(* CODESYS project PLC.project
   Title: 3D_PRINT_TITAN1
   Version: 0.0.0.0

Project tree, tasks and I/O mapping:
  Controller_2A1 : TM241CE24T/U, Schneider Electric, order no. TM241CE24T/U, version 4.0.6.18
    application Application
      libraries: SysTime, 3.4.1.20 (System)
      task MAST (cyclic, interval t#10ms, priority 1, watchdog 1000 ms x 1) calls AVC, Main
      program Main [ST]
      trace Trace_2 (task MAST): Freq_WF1, Freq_WF2, Freq_WF3
      program Wire_Speed_Correction [ST]
      program Manual [ST]
      program Auto [ST]
      trace Trace_3 (task MAST): Process_Auto, MW6, MW4
      program Alarms_manual [ST]
      program Measure [ST]
      trace Trace (task MAST): qiModule_4A1_QW0
      program Alarms_auto [ST]
      trace Trace_1 (task MAST): EM_L_PWM, EM_R_PWM
      program AVC [ST]
      global variables GVL
    Counters : Counters, Schneider Electric, version 4.0.6.18
        settings: A input History = 'old=4 new=-1'; A input History = 'old=4 new=-1'; Instance name = 'HSC0'; A input History = 'old=-1 new=4'; Temporary Instance name = 'HSC0'; Instance name = 'HSC1'; A input History = 'old=-1 new=5'; Temporary Instance name = 'HSC1'; Instance name = 'HSC2'; A input History = 'old=-1 new=6'; Temporary Instance name = 'HSC2'
    Cartridge_1 : Cartridge, Schneider Electric, version 4.0.6.18
    Serial_Line_1 : Serial line, Schneider Electric, version 4.0.6.18
      Modbus_IOScanner : Modbus IOScanner, Schneider Electric, version 3.5.3.8
          settings: Transmission = 'RTU'; ResponseTimeout = 1000; TimeBetweenFrames = 10
        Generic_Modbus_Slave : Generic Modbus Slave, Schneider Electric, version 3.5.3.9
            settings: SlaveAddress = 10; ResponseTimeout = 5000; Output.Function Code = 16; Output.Read Offset = 0; Output.Read Length = 0; Output.Write Offset = 16#0000; Output.Write Length = 1; Output.Cycle Time = 10
            unmapped channels: Output
    DI : Digital Inputs, Schneider Electric, version 4.0.6.18
        settings: IOs Usage = 112
        input  ibDI_IB1 : BYTE  // IB1
        unmapped channels: IW0
    Pulse_Generators : Pulse Generators, Schneider Electric, version 4.0.6.18
        settings: A output History = 'old=0 new=-1'; A output History = 'old=1 new=-1'; A output History = 'old=2 new=-1'
    Serial_Line_2 : Serial line, Schneider Electric, version 4.0.6.18
      Modbus_Manager : Modbus Manager, Schneider Electric, version 4.0.0.2
    DQ : Digital Outputs, Schneider Electric, version 4.0.6.18
        output qwDQ_QW0 : WORD  // QW0
        output qbDQ_QB1 : BYTE  // QB1
    COM_Bus : COM bus, Schneider Electric, version 4.0.6.18
    IO_Bus : IO bus - TM3, Schneider Electric, version 4.0.6.18
      Module_7A1 : TM3AM6/G, Schneider Electric, order no. TM3AM6/G, version 1.0.0.14
          settings: KPI Configuration.KPI Configuration[32] = 19; KPI Configuration.KPI Configuration[33] = 19; KPI Configuration.KPI Configuration[34] = 160; KPI Configuration.KPI Configuration[35] = 15; KPI Configuration.KPI Configuration[36] = 160; KPI Configuration.KPI Configuration[37] = 15; KPI Configuration.KPI Configuration[38] = 32; KPI Configuration.KPI Configuration[39] = 78; KPI Configuration.KPI Configuration[40] = 32; KPI Configuration.KPI Configuration[41] = 78
          input  iiModule_2_IW0 : INT  // IW0
          input  iiModule_2_IW1 : INT  // IW1
          input  iiModule_2_IW2 : INT  // IW2
          input  iiModule_2_IW3 : INT  // IW3
          output qiModule_2_QW0 : INT  // QW0
          output qiModule_2_QW1 : INT  // QW1
          input  ibModule_2_IBStatusIW0 : BYTE  // IBStatusIW0
          input  ibModule_2_IBStatusIW1 : BYTE  // IBStatusIW1
          input  ibModule_2_IBStatusIW2 : BYTE  // IBStatusIW2
          input  ibModule_2_IBStatusIW3 : BYTE  // IBStatusIW3
          input  ibModule_2_IBStatusQW0 : BYTE  // IBStatusQW0
          input  ibModule_2_IBStatusQW1 : BYTE  // IBStatusQW1
      Module_5A1 : TM3AQ4/G, Schneider Electric, order no. TM3AQ4/G, version 1.0.0.12
          settings: KPI Configuration.KPI Configuration[0] = 19; KPI Configuration.KPI Configuration[1] = 19; KPI Configuration.KPI Configuration[2] = 19; KPI Configuration.KPI Configuration[3] = 19; KPI Configuration.KPI Configuration[4] = 160; KPI Configuration.KPI Configuration[5] = 15; KPI Configuration.KPI Configuration[6] = 160; KPI Configuration.KPI Configuration[7] = 15; KPI Configuration.KPI Configuration[8] = 160; KPI Configuration.KPI Configuration[9] = 15; KPI Configuration.KPI Configuration[10] = 160; KPI Configuration.KPI Configuration[11] = 15; KPI Configuration.KPI Configuration[12] = 32; KPI Configuration.KPI Configuration[13] = 78; KPI Configuration.KPI Configuration[14] = 32; KPI Configuration.KPI Configuration[15] = 78; KPI Configuration.KPI Configuration[16] = 32; KPI Configuration.KPI Configuration[17] = 78; KPI Configuration.KPI Configuration[18] = 32; KPI Configuration.KPI Configuration[19] = 78
          output qiModule_5A1_QW0 : INT  // QW0
          output qiModule_5A1_QW1 : INT  // QW1
          output qiModule_5A1_QW2 : INT  // QW2
          output qiModule_5A1_QW3 : INT  // QW3
          input  ibModule_5A1_IBStatusQW0 : BYTE  // IBStatusQW0
          input  ibModule_5A1_IBStatusQW1 : BYTE  // IBStatusQW1
          input  ibModule_5A1_IBStatusQW2 : BYTE  // IBStatusQW2
          input  ibModule_5A1_IBStatusQW3 : BYTE  // IBStatusQW3
      Module_9A1 : TM3TI4/G, Schneider Electric, order no. TM3TI4/G, version 1.0.1.5
          settings: KPI Configuration.KPI Configuration[1] = 35; KPI Configuration.KPI Configuration[2] = 35; KPI Configuration.KPI Configuration[7] = 0; KPI Configuration.KPI Configuration[8] = 160; KPI Configuration.KPI Configuration[9] = 15; KPI Configuration.KPI Configuration[14] = 48; KPI Configuration.KPI Configuration[15] = 117; KPI Configuration.KPI Configuration[16] = 32; KPI Configuration.KPI Configuration[17] = 78; KPI Configuration.KPI Configuration[22] = 5; KPI Configuration.KPI Configuration[24] = 10
          input  iiModule_3_IW0 : INT  // IW0
          input  iiModule_3_IW1 : INT  // IW1
          input  iiModule_3_IW2 : INT  // IW2
          input  iiModule_3_IW3 : INT  // IW3
          input  ibModule_3_IBStatusIW0 : BYTE  // IBStatusIW0
          input  ibModule_3_IBStatusIW1 : BYTE  // IBStatusIW1
          input  ibModule_3_IBStatusIW2 : BYTE  // IBStatusIW2
          input  ibModule_3_IBStatusIW3 : BYTE  // IBStatusIW3
      Module_3A1 : TM3DQ8T/G, Schneider Electric, order no. TM3DQ8T/G, version 1.0.1.4
          output qbModule_1_QB0 : BYTE  // QB0
      Module_3A2 : TM3DQ16R/G, Schneider Electric, order no. TM3DQ16R/G, version 1.0.1.4
          output qwModule_1_QW0 : WORD  // QW0
      Module_4A1 : TM3AQ4/G, Schneider Electric, order no. TM3AQ4/G, version 1.0.0.12
          settings: KPI Configuration.KPI Configuration[0] = 19; KPI Configuration.KPI Configuration[1] = 19; KPI Configuration.KPI Configuration[2] = 19; KPI Configuration.KPI Configuration[3] = 19; KPI Configuration.KPI Configuration[4] = 160; KPI Configuration.KPI Configuration[5] = 15; KPI Configuration.KPI Configuration[6] = 160; KPI Configuration.KPI Configuration[7] = 15; KPI Configuration.KPI Configuration[8] = 160; KPI Configuration.KPI Configuration[9] = 15; KPI Configuration.KPI Configuration[10] = 160; KPI Configuration.KPI Configuration[11] = 15; KPI Configuration.KPI Configuration[12] = 32; KPI Configuration.KPI Configuration[13] = 78; KPI Configuration.KPI Configuration[14] = 32; KPI Configuration.KPI Configuration[15] = 78; KPI Configuration.KPI Configuration[16] = 32; KPI Configuration.KPI Configuration[17] = 78; KPI Configuration.KPI Configuration[18] = 32; KPI Configuration.KPI Configuration[19] = 78
          output qiModule_4A1_QW0 : INT  // QW0
          output qiModule_4A1_QW1 : INT  // QW1
          output qiModule_4A1_QW2 : INT  // QW2
          output qiModule_4A1_QW3 : INT  // QW3
          input  ibModule_4A1_IBStatusQW0 : BYTE  // IBStatusQW0
          input  ibModule_4A1_IBStatusQW1 : BYTE  // IBStatusQW1
          input  ibModule_4A1_IBStatusQW2 : BYTE  // IBStatusQW2
          input  ibModule_4A1_IBStatusQW3 : BYTE  // IBStatusQW3
    Ethernet_Slave : Ethernet Network, Schneider Electric, version 4.0.6.18
        settings: IPAddress = [192, 168, 137, 2]; SubnetMask = [255, 255, 255, 0]; DeviceName = 'PLC_Slave'; WebServer = FALSE; FTP Server = FALSE; SoMachine Protocol = TRUE; Modbus Server = TRUE; NetManage Protocol = FALSE; SNMP protocol = FALSE
  FdtConnections : FDT Connections, Schneider Electric, version 1.0.0.2
    Modbus_Serial_Line_Manager : Modbus Serial Line Manager, Schneider Electric, version 2.2.5
*)

// Controller_2A1/Application/GVL
VAR_GLOBAL
	IX07 AT %IX0.7: BOOL;
	IW19 AT %IW19: WORD ;
	QW13 AT %QW13: WORD;
    Robot_MeasureCmd : BOOL; // 1 = міряти, 0 = зупинити
    Robot_MeasureCmd_Prev : BOOL := FALSE; // Попередній стан сигналу
    // Події
    StartEvent : BOOL := FALSE;
    StopEvent : BOOL := FALSE;
    // Стан вимірювання
    Measuring : BOOL := FALSE;
    MeasureDone : BOOL := FALSE;
    MeasureStatus : INT := 0;     // 0=idle, 1=measuring, 2=done, 3=error
    // Аналоговий сигнал
    VoltageRaw : REAL;
    VoltageFiltered : REAL;
    // Фільтрація
    K_Filter : REAL := 0.12;
    FirstSample : BOOL := TRUE;
    // Обмеження допустимого діапазону
    VoltageMin : REAL := 10.0;
    VoltageMax : REAL := 30.0;
    // Захист від різких викидів
    MaxJump : REAL := 10.0;
    SampleValid : BOOL := FALSE;
    // Накопичення середнього
    VoltageSum : REAL := 0.0;
    SampleCount : DINT := 0;
    VoltageAverage : REAL := 0.0;
    // Результат для Modbus
    VoltageAverage_x100 : WORD := 0;
	
	AVC_ON: BOOL;	
	AVC_Correction AT %QW13: UINT;
	PilotArcIN AT %IX0.0: BOOL;
	PilotArc: BOOL;
	MainArc AT %IX0.1: BOOL;
	//EncoderWF1 AT %IX0.4: BOOL;
	//EncoderWF2 AT %IX0.5: BOOL;
	//EncoderWF3 AT %IX0.6: BOOL;
	StartExt AT %IX1.0: BOOL;
	ReadyExt AT %IX1.1: BOOL;
	EmergencyExt AT %IX1.2: BOOL;
	
	EM_R_PWM AT %QX0.0: BOOL;
	EM_L_PWM AT %QX0.1: BOOL;
	EM_R_EN AT %QX0.2: BOOL;
	EM_L_EN AT %QX0.3: BOOL;
	StartParc AT %QX0.4: BOOL;
	StartMArc AT %QX0.5: BOOL;
	PArcON AT %QX0.6: BOOL;
	ProcON AT %QX0.7: BOOL;
	
	MF1_CW AT %QX3.0: BOOL;
	MF1_CCW AT %QX3.1: BOOL;
	MF2_CW AT %QX3.2: BOOL;
	MF2_CCW AT %QX3.3: BOOL;
	MF3_CW AT %QX3.4: BOOL;
	MF3_CCW AT %QX3.5: BOOL;
	
	Y1 AT %QX4.0: BOOL;
	Y2 AT %QX4.1: BOOL;
	Y3 AT %QX4.2: BOOL;
	Y4 AT %QX4.3: BOOL;
	Y5 AT %QX4.4: BOOL;
	Y6 AT %QX4.5: BOOL;
	Y7 AT %QX4.6: BOOL;
	Y8 AT %QX4.7: BOOL;
	
	PF1 AT %QX5.0: BOOL;
	PF2 AT %QX5.1: BOOL;
	PF3 AT %QX5.2: BOOL;
	PF4 AT %QX5.3: BOOL;
	
	CMT_PS AT %QX5.4: BOOL;
	CMT_PlusI AT %QX5.5: BOOL;
	CMT_MinusI AT %QX5.6: BOOL;
	
	PF1_SPD AT %QW3: WORD;
	PF2_SPD AT %QW4: WORD;
	PF3_SPD AT %QW5: WORD;
	PF4_SPD AT %QW6: WORD;
	
	WF1_SPD AT %QW7: WORD;
	WF2_SPD AT %QW8: WORD;
	WF3_SPD AT %QW9: WORD;
	
	SetCurrent AT %QW11: WORD;
	MeasureU AT %IW14: WORD;
	MeasureI AT %IW15: WORD;
	MeasureU_MHI AT %MW100: WORD;
	MeasureI_MHI AT %MW102: WORD;
	Alarms AT %MW104 : WORD;
	ErrorInManual AT %MW106: WORD;
	
	EmagFreqCalc: REAL;
	Toggle_Ready : BOOL;
	ToggleState : BOOL;
	LastToggleTime : ULINT := 0;
	CurrentTime : ULINT;
    HalfPeriod_us : ULINT;
	
	
	EmagFreqCalc_Auto: REAL;

	Freq_WF1 : REAL := 0.0;
	Freq_WF2 : REAL := 0.0;
	Freq_WF3 : REAL := 0.0;
	Correction : BOOL;
	
	Enable_Start : BOOL;
	
	TON_Delay_Start_PF : TON;
	TON_Delay_Start_WF : TON;
	TON_Delay_Start_Emagnet : TON;
	TON_preblow : TON;
	
	
	MW0 AT %MW0: WORD;
	MW2 AT %MW2: WORD;
	MW4 AT %MW4 : WORD;
	MW6 AT %MW6 : WORD;
	MW8 AT %MW8 : WORD;
	PrevCurrentCMT_HMI : WORD;
END_VAR

VAR_GLOBAL RETAIN	
	EmagFreqSet AT %MD11: REAL;
	
	AVC_Voltage AT %MW12: WORD;
	AVC_Accuracy AT %MW14: WORD;
	AVC_PID_Kp AT %MD8: REAL;
	AVC_PID_Ki AT %MD55: REAL;
	AVC_DELAY AT %MW114: WORD;
	
	SetCurrent_HMI_Man AT %MW20: WORD;
	WF1_SPD_HMI_Man AT %MW26: WORD;
	WF2_SPD_HMI_Man AT %MW28: WORD;
	WF3_SPD_HMI_Man AT %MW30: WORD;
	PF1_SPD_HMI_Man AT %MW32: WORD;
	PF2_SPD_HMI_Man AT %MW34: WORD;
	PF3_SPD_HMI_Man AT %MW36: WORD;
	PF4_SPD_HMI_Man AT %MW38: WORD;
	SetCurrentCMT_HMI AT %MW40: WORD;
	Check_Voltage_Current_Delay AT %MW42 : WORD;
	Emergency_Delay AT %MW44 : WORD;
	Auto_Button_State AT %MW46 : WORD;
	Set_Emergency_Voltage AT %MW48 : WORD;
	Set_Emergency_Current AT %MW50 : WORD;
	
	EmagFreqSet_Auto AT %MD27: REAL;
	SetCurrent_HMI_Auto AT %MW52: WORD;
	WF1_SPD_HMI_Auto AT %MW58: WORD;
	WF2_SPD_HMI_Auto AT %MW60: WORD;
	WF3_SPD_HMI_Auto AT %MW62: WORD;
	PF1_SPD_HMI_Auto AT %MW64: WORD;
	PF2_SPD_HMI_Auto AT %MW66: WORD;
	PF3_SPD_HMI_Auto AT %MW68: WORD;
	PF4_SPD_HMI_Auto AT %MW70: WORD;
	Delay_Gas_Preblow AT %MW74 : WORD;
 	Delay_Gas_Finishblow AT %MW76 : WORD;
	Delay_Gas_Analysys AT %MW78 : WORD;
	Process_Auto AT %MW80 : WORD;
	Delay_Start_PF AT %MW82 : WORD;
	Delay_Start_WF AT %MW84 : WORD;
	Delay_Start_Emagnet AT %MW86 : WORD;
	Delay_Stop_PF AT %MW88 : WORD;
	Delay_Stop_WF AT %MW90 : WORD;
	Delay_Stop_Emagnet AT %MW92 : WORD;
	Delay_Analysys_Pilot AT %MW94 : WORD;
	Delay_Analysys_Main AT %MW96 : WORD;  
END_VAR

// Controller_2A1/Application/AVC
PROGRAM AVC
VAR
	PID_1: PID;
	RAMP_INT_1: RAMP_INT;
	TON_AVC: TON;
	TON_StopConfirm: TON;
	Robot_MeasureCmd_Raw: BOOL;
END_VAR

// Визначення фронтів одного дискретного сигналу
Robot_MeasureCmd := IX07;

// START: фронт 0 -> 1
StartEvent := Robot_MeasureCmd AND NOT Robot_MeasureCmd_Prev;

// STOP: фронт 1 -> 0
StopEvent := NOT Robot_MeasureCmd AND Robot_MeasureCmd_Prev;

TON_AVC(IN:= NOT Robot_MeasureCmd, PT:= T#5000MS); //Захист від надсилання старих даних
IF TON_AVC.Q THEN QW13:= 0; END_IF //Захист від надсилання старих даних

// START: сигнал від робота перейшов 0 -> 1
IF StartEvent THEN
    Measuring := TRUE; MeasureDone := FALSE; MeasureStatus := 1; VoltageSum := 0.0; SampleCount := 0; VoltageAverage := 0.0; VoltageFiltered := 0.0; FirstSample := TRUE; END_IF;

// Вимірювання, поки Robot_MeasureCmd = TRUE
IF Measuring AND Robot_MeasureCmd THEN
    VoltageRaw := WORD_TO_REAL(MeasureU) / 1000.0;
    SampleValid := (VoltageRaw >= VoltageMin) AND (VoltageRaw <= VoltageMax); // Перевірка допустимого діапазону
    IF SampleValid THEN
        IF FirstSample THEN
            VoltageFiltered := VoltageRaw;
            FirstSample := FALSE;
            VoltageSum := VoltageSum + VoltageFiltered;
            SampleCount := SampleCount + 1;
        ELSE
            IF ABS(VoltageRaw - VoltageFiltered) <= MaxJump THEN // Захист від одиночних викидів
                VoltageFiltered := VoltageFiltered + K_Filter * (VoltageRaw - VoltageFiltered); // EMA-фільтр
                VoltageSum := VoltageSum + VoltageFiltered; // Накопичення середнього по відфільтрованому сигналу
                SampleCount := SampleCount + 1;
            END_IF;
        END_IF;
    END_IF;
END_IF;

// STOP: сигнал від робота перейшов 1 -> 0
IF StopEvent THEN
    Measuring := FALSE;
    IF SampleCount > 0 THEN
        VoltageAverage := VoltageSum / DINT_TO_REAL(SampleCount); VoltageAverage_x100 := REAL_TO_WORD(VoltageAverage * 100.0); MeasureStatus := 2;
    ELSE
        VoltageAverage := 0.0; VoltageAverage_x100 := 0; MeasureStatus := 3;
    END_IF;
    MeasureDone := TRUE;
	QW13:= VoltageAverage_x100;
END_IF;

// Запам'ятовуємо попередній стан сигналу
Robot_MeasureCmd_Prev := Robot_MeasureCmd;

END_PROGRAM

// Controller_2A1/Application/Main
PROGRAM Main
VAR
	RTRIG1: R_TRIG;
END_VAR

Measure();
Wire_Speed_Correction();
RTRIG1(CLK:= TRUE); //Тригер присвоєння струму при старті
IF RTRIG1.Q THEN PrevCurrentCMT_HMI:= SetCurrentCMT_HMI; END_IF
IF MW0.0 THEN Auto(); Alarms_auto(); ELSE  Manual(); Alarms_manual(); END_IF

END_PROGRAM

// Controller_2A1/Application/Measure
PROGRAM Measure
VAR
	R_TRIG_WF1: R_TRIG;
	R_TRIG_WF3: R_TRIG;
	R_TRIG_WF2: R_TRIG;
	TON_READY_EXT: TON;
	STATE_READY_EXT: BOOL;
	ReadyExt_Prev: BOOL;
	ReadyExt_Reset: BOOL;
	PArc_trig: R_TRIG;
END_VAR

IF ReadyExt <> ReadyExt_Prev THEN ReadyExt_Reset:= FALSE; ReadyExt_Prev:= ReadyExt; ELSE  ReadyExt_Reset:= TRUE; END_IF //Обнулення лічильника Ready ext
TON_READY_EXT(IN:= ReadyExt_Reset, PT:= T#150MS, Q=> STATE_READY_EXT); //Лічильник Ready ext
MeasureU_MHI:= MeasureU;
MeasureI_MHI:= MeasureI;
MW0.1:= StartExt;
MW0.2:= NOT(STATE_READY_EXT);
MW0.3:= NOT(EmergencyExt);
MW0.4:= PilotArcIN; 
MW0.5:= MainArc;

PArc_trig(CLK:= PilotArcIN); //Тригер наявності черг дуг
IF PArc_trig.Q THEN PilotArc:= TRUE; END_IF //Взведення флажка черг дуг
IF NOT(StartParc) THEN PilotArc:= FALSE; END_IF //Скидання флажка черг дуг

// Ввікмнення лічильника імпульсів
//WF1
HSC0.EN_Enable := TRUE;
HSC0.F_Enable := TRUE;
HSC0();
Freq_WF1 := DINT_TO_REAL(HSC0.CurrentValue);
//WF2
HSC1.EN_Enable := TRUE;
HSC1.F_Enable := TRUE;
HSC1();
Freq_WF2 := DINT_TO_REAL(HSC1.CurrentValue);
//WF3
HSC2.EN_Enable := TRUE;
HSC2.F_Enable := TRUE;
HSC2();
Freq_WF2 := DINT_TO_REAL(HSC2.CurrentValue);

PArcON:= PilotArc; //Pilot arc ON for robot

END_PROGRAM

// Controller_2A1/Application/Wire_Speed_Correction
PROGRAM Wire_Speed_Correction
VAR
	New_WF1_SPD: WORD;
	LastCorrTime: ULINT := 0;
	TimeDiff: TIME;
	CurrentTime_WF: ULINT;
	LastTime_WF: ULINT := 0;
	Wanted_Speed_WF1: REAL;
	Wanted_Speed_WF2: REAL;
	Wanted_Speed_WF3: REAL;
	HMI_Old_WF1: WORD;
	HMI_Old_WF2: WORD;
	New_WF2_SPD: WORD;
	HMI_Old_WF3: WORD;
	New_WF3_SPD: WORD;
END_VAR

// Отримання поточного часу в мікросекундах
SysTimeGetUs(CurrentTime_WF);

// Розрахунок бажаної швидкості в імпульсах
IF MW0.0 THEN
	Wanted_Speed_WF1 := (WORD_TO_REAL(WF1_SPD_HMI_Auto) - 6000.0) * ((1700.0-100.0) / (20000.0-6000.0)) + 100.0;
	Wanted_Speed_WF2 := (WORD_TO_REAL(WF2_SPD_HMI_Auto) - 6000.0) * ((1700.0-100.0) / (20000.0-6000.0)) + 100.0;
	Wanted_Speed_WF3 := (WORD_TO_REAL(WF3_SPD_HMI_Auto) - 6000.0) * ((1700.0-100.0) / (20000.0-6000.0)) + 100.0;
			// Ініціалізація
	IF HMI_Old_WF1 <> WF1_SPD_HMI_Auto AND MW4.12 AND Process_Auto = 3 THEN HMI_Old_WF1 := WF1_SPD_HMI_Auto; New_WF1_SPD := HMI_Old_WF1; END_IF
	IF HMI_Old_WF2 <> WF2_SPD_HMI_Auto AND MW4.13 AND Process_Auto = 3 THEN HMI_Old_WF2 := WF2_SPD_HMI_Auto; New_WF2_SPD := HMI_Old_WF2; END_IF
	IF HMI_Old_WF3 <> WF3_SPD_HMI_Auto AND MW4.14 AND Process_Auto = 3 THEN HMI_Old_WF3 := WF3_SPD_HMI_Auto; New_WF3_SPD := HMI_Old_WF3; END_IF
ELSE
	Wanted_Speed_WF1 := (WORD_TO_REAL(WF1_SPD_HMI_Man) - 6000.0) * ((1700.0-100.0) / (20000.0-6000.0)) + 100.0;
	Wanted_Speed_WF2 := (WORD_TO_REAL(WF2_SPD_HMI_Man) - 6000.0) * ((1700.0-100.0) / (20000.0-6000.0)) + 100.0;
	Wanted_Speed_WF3 := (WORD_TO_REAL(WF3_SPD_HMI_Man) - 6000.0) * ((1700.0-100.0) / (20000.0-6000.0)) + 100.0;
		// Ініціалізація
	IF HMI_Old_WF1 <> WF1_SPD_HMI_Man AND MW2.04 THEN HMI_Old_WF1 := WF1_SPD_HMI_Man; New_WF1_SPD := HMI_Old_WF1; END_IF
	IF HMI_Old_WF2 <> WF2_SPD_HMI_Man AND MW2.06 THEN HMI_Old_WF2 := WF2_SPD_HMI_Man; New_WF2_SPD := HMI_Old_WF2; END_IF
	IF HMI_Old_WF3 <> WF3_SPD_HMI_Man AND MW2.08 THEN HMI_Old_WF3 := WF3_SPD_HMI_Man; New_WF3_SPD := HMI_Old_WF3; END_IF
END_IF


// Обчислення раз на секунду
	IF (CurrentTime_WF - LastTime_WF) >= REAL_TO_ULINT(100_000.0) THEN
		//WF1
		IF MW2.04 OR (MW4.12 AND Process_Auto = 3) THEN
		 	IF Wanted_Speed_WF1 - Freq_WF1 > 5.0 THEN New_WF1_SPD := New_WF1_SPD + 37; ELSIF Freq_WF1 - Wanted_Speed_WF1 > 5.0 THEN New_WF1_SPD := New_WF1_SPD - 37; END_IF
			 	LastTime_WF := CurrentTime_WF; // обнулення таймера
		END_IF
		//WF2
   		IF MW2.06 OR (MW4.13 AND Process_Auto = 3) THEN
		 	IF Wanted_Speed_WF2 - Freq_WF2 > 5.0 THEN New_WF2_SPD := New_WF2_SPD + 37; ELSIF Freq_WF2 - Wanted_Speed_WF2 > 5.0 THEN New_WF2_SPD := New_WF2_SPD - 37; END_IF
			 	LastTime_WF := CurrentTime_WF; // обнулення таймера
		END_IF
		//WF3
		IF MW2.08 OR (MW4.14 AND Process_Auto = 3) THEN
		 	IF Wanted_Speed_WF3 - Freq_WF3 > 5.0 THEN New_WF3_SPD := New_WF3_SPD + 37; ELSIF Freq_WF3 - Wanted_Speed_WF3 > 5.0 THEN New_WF3_SPD := New_WF3_SPD - 37; END_IF
			 	LastTime_WF := CurrentTime_WF; // обнулення таймера
		END_IF
	END_IF


// Обмеження діапазону напруги
IF New_WF1_SPD > 20000 THEN New_WF1_SPD := 20000; ELSIF New_WF1_SPD < 6000 THEN New_WF1_SPD := 6000; END_IF
IF New_WF2_SPD > 20000 THEN New_WF2_SPD := 20000; ELSIF New_WF2_SPD < 6000 THEN New_WF2_SPD := 6000; END_IF
IF New_WF3_SPD > 20000 THEN New_WF3_SPD := 20000; ELSIF New_WF3_SPD < 6000 THEN New_WF3_SPD := 6000; END_IF

// Встановлення остаточного значення
WF1_SPD := NEW_WF1_SPD;
WF2_SPD := NEW_WF2_SPD;
WF3_SPD := NEW_WF3_SPD;

END_PROGRAM

// Controller_2A1/Application/Auto
PROGRAM Auto
VAR
	TON_After_Stop: TON;
	TON_After_Stop_state: BOOL;
	TON_Finish_blow: TON;
	TON_Finish_blow_state: BOOL;
	TON_CMT: TON;
	TON_CMT_State: BOOL;
	TON_CMT1: TON;
	TON_CMT_State1: BOOL;
	Counter: INT;
	R_TRIG_state: BOOL;
	Prev_MW4_15: BOOL;
	Prev_MW6_0: BOOL;
	TON_Delay_Stop_PF: TON;
	TON_Delay_Stop_WF: TON;
	TON_Delay_Stop_Emagnet: TON;
	R_TRIG_External: R_TRIG;
	TON_Alarm: TON;
	TON_Alarm2: TON;
	Step: BOOL;
	Allow_finish_blow: BOOL;
	Prev_Process: WORD;
END_VAR

// Встановлення Powder Feeder
IF MW4.7 THEN PF1_SPD := PF1_SPD_HMI_Auto; END_IF
IF MW4.8 THEN PF2_SPD := PF2_SPD_HMI_Auto; END_IF
IF MW4.9 THEN PF3_SPD := PF3_SPD_HMI_Auto; END_IF
IF MW4.10 THEN PF4_SPD := PF4_SPD_HMI_Auto; END_IF

// E-magnet
IF MW4.11 THEN 
	IF EmagFreqSet_Auto > 0 THEN EmagFreqCalc_Auto:= EmagFreqSet_Auto; ELSE EmagFreqCalc_Auto:= 10; END_IF //Обхід помилки ділення на нуль для прорахунку частоти ел.маг.
END_IF

// Встановлення Wire Feeder
IF MW4.12 THEN WF1_SPD := WF1_SPD_HMI_Auto; END_IF
IF MW4.13 THEN WF2_SPD := WF2_SPD_HMI_Auto; END_IF
IF MW4.14 THEN WF3_SPD := WF3_SPD_HMI_Auto; END_IF


// Ввімкнення іншого режиму
IF MW6.0 AND NOT Prev_MW6_0 AND Auto_Button_State = 0 THEN 
	MW4.7 := FALSE; MW4.8 := FALSE; MW4.9 := FALSE; MW4.10 := FALSE; MW4.11 := FALSE; MW4.15 := FALSE;
END_IF
IF MW4.15 AND NOT Prev_MW4_15 AND Auto_Button_State = 0 THEN 
	MW6.0 := FALSE; 
END_IF
IF Auto_Button_State = 0 THEN Prev_MW6_0 := MW6.0; Prev_MW4_15 := MW4.15; ELSE MW6.0 :=  Prev_MW6_0;  MW4.15:=Prev_MW4_15; END_IF
 

// Якщо CMT
IF MW6.0 THEN 
	MW4.7 := FALSE; MW4.8 := FALSE; MW4.9 := FALSE; MW4.10 := FALSE; MW4.11 := FALSE;
END_IF


IF Step = FALSE THEN
    TON_Alarm(IN := TRUE, PT := T#500MS);
    TON_Alarm2(IN := FALSE);
ELSE
    TON_Alarm2(IN := TRUE, PT := T#500MS);
    TON_Alarm(IN := FALSE);
END_IF;


// Alarm
IF (MW6.10 OR NOT(EmergencyExt)) AND Process_Auto <> 0 AND Auto_Button_State = 0 AND Alarms <> 0 THEN
	IF TON_Alarm.Q THEN
    	Process_Auto := 10;
    	Step := TRUE; 
    	TON_Alarm(IN := FALSE);
	END_IF;
	IF TON_Alarm2.Q THEN
    	Process_Auto := 11;
    	Step := FALSE; 
    	TON_Alarm2(IN := FALSE); 
	END_IF;
	MW6.9 := FALSE;
	Enable_Start := FALSE; 
	TON_Delay_Start_PF(IN:=FALSE); TON_Delay_Start_Emagnet(IN:=FALSE); TON_Delay_Start_WF(IN:=FALSE);TON_preblow(IN:=FALSE);
ELSIF NOT(MW6.11) AND Auto_Button_State = 0 THEN 
	Process_Auto := 5; 
	MW6.9 := FALSE;
	Enable_Start := FALSE;
END_IF

// Блок старту
IF NOT(MW4.3) AND Process_Auto <> 5 AND MW6.11 OR Enable_Start THEN MW6.6 := FALSE; ELSE MW6.6 := TRUE; END_IF

//Зовнішній пуск
R_TRIG_External(CLK:=StartExt);

// Local start
IF NOT(MW4.3) AND MW6.11 AND (MW6.5 AND Auto_Button_State = 0) THEN 
	IF NOT(Enable_Start) THEN
		//Are you sure
			MW6.9 := TRUE;
		Enable_Start := TRUE;
	END_IF
ELSIF MW4.3 AND R_TRIG_External.Q AND MW6.11 THEN// External start
	IF NOT(Enable_Start) THEN MW6.12 := TRUE; END_IF
	Enable_Start := TRUE;
	MW6.5 := TRUE;
END_IF
//Close are you sure
IF MW2.15 OR MW4.3 OR (NOT(MW6.11) AND Auto_Button_State = 0) OR (NOT(EmergencyExt) AND Auto_Button_State = 0) THEN Enable_Start := FALSE; MW6.9 := FALSE; MW2.15 := FALSE; MW6.5 := FALSE; END_IF

//Set process to ready
IF NOT(Enable_Start) AND MW6.11 AND Auto_Button_State = 0 THEN Process_Auto := 0; END_IF


// Start Process
IF MW6.12 AND Enable_Start AND MW6.11 THEN
	
	//Block Manual
	MW6.13 := TRUE;
	
	//Block Start
	MW6.6 := FALSE;
	
	//Close Are you sure
	MW6.9 := FALSE;
	
	//Process ON
	Auto_Button_State := 1;
	
	//Preblow
	IF Y1 AND NOT(Y2) AND NOT(Y3) AND NOT(Y4) THEN Y1 := TRUE; MW6.1:= TRUE; ELSE Y1 := MW6.1; END_IF
	IF NOT(Y1) AND Y2 AND NOT(Y3) AND NOT(Y4) THEN Y2 := TRUE; MW6.2:= TRUE;ELSE Y2 := MW6.2; END_IF
	IF NOT(Y1) AND NOT(Y2) AND Y3 AND NOT(Y4) THEN Y3 := TRUE; MW6.3:= TRUE;ELSE Y3 := MW6.3; END_IF
	IF NOT(Y1) AND NOT(Y2) AND NOT(Y3) AND Y4 THEN Y4 := TRUE; MW6.4:= TRUE;ELSE Y4 := MW6.4; END_IF
		
	IF NOT(TON_preblow.Q) THEN Process_Auto := 1; END_IF
	
	TON_preblow(IN:=Enable_Start , PT:=WORD_TO_TIME(Delay_Gas_Preblow));
	//PLASMA
	IF MW4.15 THEN 
		SetCurrent:= SetCurrent_HMI_Auto; //Current set
		//Pilot Arc
		IF TON_preblow.Q AND MW6.11 THEN 
			StartParc:= TRUE; 
			IF NOT(PilotArc) THEN Process_Auto := 2; END_IF 
		END_IF
		//Main Arc
		IF PilotArc AND StartParc THEN 
			StartMArc:= TRUE; 
			IF NOT(MainArc) THEN Process_Auto := 8; END_IF 
		END_IF
		//Additional equipment
		IF MainArc AND Process_Auto <> 3 AND StartMArc THEN Process_Auto := 9; END_IF	
		
		//Delays
		TON_Delay_Start_PF(IN:=MainArc AND StartParc AND StartMArc AND PilotArc, PT:=WORD_TO_TIME(Delay_Start_PF));
		TON_Delay_Start_WF(IN:=MainArc AND StartParc AND StartMArc AND PilotArc, PT:=WORD_TO_TIME(Delay_Start_WF));
		TON_Delay_Start_Emagnet(IN:=MainArc AND StartParc AND StartMArc AND PilotArc, PT:=WORD_TO_TIME(Delay_Start_Emagnet));
		
		IF TON_Delay_Start_PF.Q THEN
			// Transport Gases
			Y5 := MW4.7; Y6 := MW4.8; Y7 := MW4.9; Y8 := MW4.10;
			//Powder Feeder 
			PF1 := MW4.7; PF2 := MW4.8; PF3 := MW4.9; PF4 := MW4.10; 
		END_IF
		
		//Wire Feeder
		IF TON_Delay_Start_WF.Q THEN 
			IF MW4.12 THEN MF1_CW:= TRUE; MF1_CCW := FALSE; ELSE MF1_CW:= FALSE; MF1_CCW := FALSE;  END_IF
			IF MW4.13 THEN MF2_CW:= TRUE; MF2_CCW := FALSE; ELSE MF2_CW:= FALSE; MF2_CCW := FALSE;  END_IF
			IF MW4.14 THEN MF3_CW:= TRUE; MF3_CCW := FALSE; ELSE MF3_CW:= FALSE; MF3_CCW := FALSE;  END_IF
		END_IF
		
		//E-magnet
		IF TON_Delay_Start_Emagnet.Q THEN
			IF MW4.11 THEN
				EM_R_EN := TRUE;
				EM_L_EN := TRUE;
				HalfPeriod_us := REAL_TO_ULINT(1000000.0 / EmagFreqCalc_Auto / 2.0); //Період в мікросекундах
				SysTimeGetUs(CurrentTime); // CurrentTime ULINT
				IF (CurrentTime - LastToggleTime) >= HalfPeriod_us THEN //Перевірка пройденого часу
					ToggleState := NOT(ToggleState); //Інверсія
					LastToggleTime := CurrentTime; //Обнулення таймеру
				END_IF	
				EM_R_PWM := ToggleState;
				EM_L_PWM := NOT(ToggleState);
			ELSE
				EM_R_EN := FALSE;
				EM_L_EN := FALSE;
				EM_R_PWM := FALSE;
				EM_L_PWM := FALSE;
				ToggleState := FALSE;
				LastToggleTime := 0;
			END_IF
		END_IF
		
		//Process
		IF (
			(NOT(MW4.7 OR MW4.8 OR MW4.9 OR MW4.10) OR TON_Delay_Start_PF.Q) AND
			(NOT(MW4.12 OR MW4.13 OR MW4.14) OR TON_Delay_Start_WF.Q) AND
			(NOT(MW4.11) OR TON_Delay_Start_Emagnet.Q) AND
			TON_preblow.Q AND PilotArc AND MainArc
			) THEN
				Process_Auto := 3;
		END_IF

	// CMT 
	ELSIF MW6.0 AND Enable_Start AND TON_preblow.Q AND MW6.11 THEN
		CMT_PS := TRUE;
		IF Process_Auto <> 9 THEN IF Process_Auto <> 3 THEN Process_Auto := 9; END_IF END_IF
		//Wire Feeder
		TON_Delay_Start_WF(IN:=TON_preblow.Q, PT:=WORD_TO_TIME(Delay_Start_WF));
		IF TON_Delay_Start_WF.Q THEN
			IF MW4.12 THEN MF1_CW:= TRUE; MF1_CCW := FALSE; ELSE MF1_CW:= FALSE; MF1_CCW := FALSE;  END_IF
			IF MW4.13 THEN MF2_CW:= TRUE; MF2_CCW := FALSE; ELSE MF2_CW:= FALSE; MF2_CCW := FALSE;  END_IF
			IF MW4.14 THEN MF3_CW:= TRUE; MF3_CCW := FALSE; ELSE MF3_CW:= FALSE; MF3_CCW := FALSE;  END_IF
		END_IF
		IF NOT(MW4.12 OR MW4.13 OR MW4.14) OR TON_Delay_Start_WF.Q THEN
			Process_Auto := 3;
		END_IF
	END_IF
END_IF
	

//CMT Process
TON_CMT(IN:= CMT_PlusI OR CMT_MinusI, PT:= T#100MS, Q=> TON_CMT_State); //Таймер імпульсу для зміни значення
TON_CMT1(IN:= NOT(CMT_PlusI) AND NOT(CMT_MinusI), PT:= T#100MS, Q=> TON_CMT_State1); //Таймер паузи для зміни значення
IF SetCurrentCMT_HMI <> PrevCurrentCMT_HMI THEN 
	Counter:= WORD_TO_INT(SetCurrentCMT_HMI) -  WORD_TO_INT(PrevCurrentCMT_HMI); //рахуємо кількість імпульсів
	IF Counter > 0 THEN  //Якщо потрібно збільшувати струм
		IF TON_CMT_State1 THEN CMT_PlusI:= TRUE; END_IF //Імпульс
		IF TON_CMT_State THEN CMT_PlusI:= FALSE; PrevCurrentCMT_HMI:= PrevCurrentCMT_HMI +1; Counter:= Counter -1; END_IF //Пауза + інкремент
	ELSIF Counter < 0 THEN  //Якщо потрібно зменшувати струм
		IF TON_CMT_State1 THEN CMT_MinusI:= TRUE; END_IF  //Імпульс
		IF TON_CMT_State THEN CMT_MinusI:= FALSE; PrevCurrentCMT_HMI:= PrevCurrentCMT_HMI -1; Counter:= Counter +1; END_IF //Пауза + декремент
	END_IF
ELSE CMT_PlusI:= FALSE; CMT_MinusI:= FALSE; END_IF //Вимкнення інкрементального та декрементального реле по дефолту
		
//Stop
IF Process_Auto <> 0 AND Enable_Start AND ((MW4.3 AND NOT(StartExt)) AND EmergencyExt AND MW6.11 OR (NOT(MW6.5) AND Auto_Button_State = 1)) OR Auto_Button_State = 2 THEN // STOP
	//YES
	MW6.12 := FALSE;
	
	//Block start
	MW6.6 := TRUE;
	
	//Set stop to button
	IF Auto_Button_State <> 0 THEN Auto_Button_State := 2; END_IF
	
	//Save stop process
	IF Process_Auto <> 6 AND Process_Auto <> 4 THEN Prev_Process := Process_Auto; END_IF
	
	//Pre-blowing
	IF Prev_Process = 1 THEN
		Allow_finish_blow := TRUE;
		
	//Waiting Pilot Arc
	ELSIF Prev_Process = 2 THEN
		//Turn off Pilot Arc
		StartParc:= FALSE;
		Allow_finish_blow := TRUE;
		
	//Working Process and CMT Start
	ELSIF Prev_Process = 3 THEN
		// CMT OFF
		CMT_PS := FALSE;
		CMT_PlusI:= FALSE; CMT_MinusI:= FALSE;
		//Turn off Main Arc
		StartMArc:= FALSE;	
		//Turn off Pilot Arc
		StartParc:= FALSE;
		TON_Delay_Stop_PF(IN:=TON_Delay_Start_PF.Q, PT:=WORD_TO_TIME(Delay_Stop_PF));
		TON_Delay_Stop_WF(IN:=TON_Delay_Start_WF.Q, PT:=WORD_TO_TIME(Delay_Stop_WF));
		TON_Delay_Stop_Emagnet(IN:=TON_Delay_Start_Emagnet.Q, PT:=WORD_TO_TIME(Delay_Stop_Emagnet));
		IF (
			(NOT(MW4.7 OR MW4.8 OR MW4.9 OR MW4.10) OR (((MW4.7 OR MW4.8 OR MW4.9 OR MW4.10) AND NOT(TON_Delay_Start_PF.Q)) OR TON_Delay_Stop_PF.Q)) AND
			(NOT(MW4.12 OR MW4.13 OR MW4.14) OR (((MW4.12 OR MW4.13 OR MW4.14) AND NOT(TON_Delay_Start_WF.Q)) OR TON_Delay_Stop_WF.Q))AND
			(NOT(MW4.11) OR ((MW4.11 AND NOT(TON_Delay_Start_Emagnet.Q)) OR TON_Delay_Stop_Emagnet.Q)) 
			) THEN
				Allow_finish_blow := TRUE;
		ELSE
			Process_Auto := 6;
		END_IF
		
	//Waiting Main Arc
	ELSIF Prev_Process = 8 THEN
		//Turn off Main Arc
		StartMArc:= FALSE;
		//Turn off Pilot Arc
		StartParc:= FALSE;
		Allow_finish_blow := TRUE;
		
	//Waiting Additional equipment
	ELSIF Prev_Process = 9 THEN
		// CMT OFF
		CMT_PS := FALSE;
		CMT_PlusI:= FALSE; CMT_MinusI:= FALSE;
		//Turn off Main Arc
		StartMArc:= FALSE;	
		//Turn off Pilot Arc
		StartParc:= FALSE;
		TON_Delay_Stop_PF(IN:=TON_Delay_Start_PF.Q, PT:=WORD_TO_TIME(Delay_Stop_PF));
		TON_Delay_Stop_WF(IN:=TON_Delay_Start_WF.Q, PT:=WORD_TO_TIME(Delay_Stop_WF));
		TON_Delay_Stop_Emagnet(IN:=TON_Delay_Start_Emagnet.Q, PT:=WORD_TO_TIME(Delay_Stop_Emagnet));
		IF (
			(NOT(MW4.7 OR MW4.8 OR MW4.9 OR MW4.10) OR (((MW4.7 OR MW4.8 OR MW4.9 OR MW4.10) AND NOT(TON_Delay_Start_PF.Q)) OR TON_Delay_Stop_PF.Q) )AND
			(NOT(MW4.12 OR MW4.13 OR MW4.14) OR (((MW4.12 OR MW4.13 OR MW4.14) AND NOT(TON_Delay_Start_WF.Q)) OR TON_Delay_Stop_WF.Q))AND
			(NOT(MW4.11) OR ((MW4.11 AND NOT(TON_Delay_Start_Emagnet.Q)) OR TON_Delay_Stop_Emagnet.Q)) 
			) THEN
				Allow_finish_blow := TRUE;
		ELSE
			Process_Auto := 6;
		END_IF
	END_IF
	
	IF TON_Delay_Stop_PF.Q THEN PF1 := FALSE; PF2 := FALSE; PF3 := FALSE; PF4 := FALSE; Y5 := FALSE; Y6 := FALSE; Y7 := FALSE; Y8 := FALSE; END_IF
	IF TON_Delay_Stop_WF.Q THEN MF1_CW:= FALSE; MF1_CCW := FALSE; MF2_CW:= FALSE; MF2_CCW := FALSE; MF3_CW:= FALSE; MF3_CCW := FALSE; END_IF
	IF (MW4.11 AND NOT(TON_Delay_Start_Emagnet.Q)) OR TON_Delay_Stop_Emagnet.Q OR Allow_finish_blow THEN 
		//Вимикаємо магніт
		EM_R_EN := FALSE;
		EM_L_EN := FALSE;
		EM_R_PWM := FALSE;
		EM_L_PWM := FALSE;
		ToggleState := FALSE;
		LastToggleTime := 0;
	ELSIF Prev_Process <> 1 AND Prev_Process <> 2 AND Prev_Process <> 8 AND Auto_Button_State <> 0 THEN
		IF MW4.11 THEN
				EM_R_EN := TRUE;
				EM_L_EN := TRUE;
				HalfPeriod_us := REAL_TO_ULINT(1000000.0 / EmagFreqCalc_Auto / 2.0); //Період в мікросекундах
				SysTimeGetUs(CurrentTime); // CurrentTime ULINT
				IF (CurrentTime - LastToggleTime) >= HalfPeriod_us THEN //Перевірка пройденого часу
					ToggleState := NOT(ToggleState); //Інверсія
					LastToggleTime := CurrentTime; //Обнулення таймеру
				END_IF	
				EM_R_PWM := ToggleState;
				EM_L_PWM := NOT(ToggleState);
		END_IF
	END_IF
	//Finish blowing
	IF Allow_finish_blow THEN
				TON_Finish_blow(IN:=Enable_Start, PT:=WORD_TO_TIME(Delay_Gas_Finishblow * 10));
				//Finish blow
				IF TON_Finish_blow.Q THEN Allow_finish_blow := FALSE; Y1 := FALSE; Y2 := FALSE; Y3 := FALSE; Y4 := FALSE; Enable_Start := FALSE; Process_Auto := 0; 
				TON_Delay_Stop_PF(IN:=FALSE); TON_Delay_Stop_Emagnet(IN:=FALSE); TON_Delay_Stop_WF(IN:=FALSE); TON_Finish_blow(IN:=FALSE);
				TON_Delay_Start_PF(IN:=FALSE); TON_Delay_Start_Emagnet(IN:=FALSE); TON_Delay_Start_WF(IN:=FALSE);TON_preblow(IN:=FALSE);
				MW6.13 := FALSE;
				Auto_Button_State := 0;
				Prev_Process := 0;
				ELSE Process_Auto := 4; END_IF
	END_IF
END_IF

IF Process_Auto = 3  THEN ProcON:= TRUE; ELSE ProcON:= FALSE; END_IF //Видача ProcON на робот

//Block local control	
IF Auto_Button_State <> 0 THEN MW8.0 := TRUE; ELSE MW8.0:= FALSE; END_IF

END_PROGRAM

// Controller_2A1/Application/Manual
PROGRAM Manual
VAR
	TON0: TON;
	TON0_State: BOOL;
	TON1: TON;
	TON1_State: BOOL;
	TON2: TON;
	TON3: TON;
	TON4: TON;
	TON5: TON;
	TON2_State: BOOL;
	TON3_State: BOOL;
	TON4_State: BOOL;
	TON5_State: BOOL;
	TON_Freq: TON;
	HalfPeriod: TIME;
	HalfPeriod_time: TIME;
	TON_CMT1: TON;
	TON_CMT: TON;
	TON_CMT_State1: BOOL;
	TON_CMT_State: BOOL;
	Counter: INT;
	RTRIG_CMT: R_TRIG;
END_VAR

Y1 := MW0.8; Y2 := MW0.9; Y3 := MW0.10; Y4 := MW0.11; Y5 := MW0.12; Y6 := MW0.13; Y7 := MW0.14; Y8 := MW0.15; //Gases
//E-Magnet//
IF EmagFreqSet > 0 THEN EmagFreqCalc:= EmagFreqSet; ELSE EmagFreqCalc:= 10; END_IF //Обхід помилки ділення на нуль для прорахунку частоти ел.маг.
IF MW2.02 THEN
	EM_R_EN := TRUE;
	EM_L_EN := TRUE;
	HalfPeriod_us := REAL_TO_ULINT(1000000.0 / EmagFreqCalc / 2.0); //Період в мікросекундах
	SysTimeGetUs(CurrentTime); // CurrentTime ULINT
	IF (CurrentTime - LastToggleTime) >= HalfPeriod_us THEN //Перевірка пройденого часу
		ToggleState := NOT(ToggleState); //Інверсія
		LastToggleTime := CurrentTime; //Обнулення таймеру
	END_IF	
	EM_R_PWM := ToggleState;
	EM_L_PWM := NOT(ToggleState);
ELSE
	EM_R_EN := FALSE;
	EM_L_EN := FALSE;
	EM_R_PWM := FALSE;
	EM_L_PWM := FALSE;
	ToggleState := FALSE;
	LastToggleTime := 0;
END_IF
//E-Magnet//
PF1:= MW2.10; PF2:= MW2.11; PF3:= MW2.12; PF4:= MW2.13; //Powder feeders
PF1_SPD:= PF1_SPD_HMI_Man; PF2_SPD:= PF2_SPD_HMI_Man; PF3_SPD:= PF3_SPD_HMI_Man; PF4_SPD:= PF4_SPD_HMI_Man; //Powder feeders speed
//Wire feeders//
TON0(IN:= MW2.5, PT:= T#1MS, Q=> TON0_State); //Set1 dir1
TON1(IN:= NOT(MW2.5), PT:= T#1MS, Q=> TON1_State); //Set1 dir2
TON2(IN:= MW2.7, PT:= T#1MS, Q=> TON2_State); //Set2 dir1
TON3(IN:= NOT(MW2.7), PT:= T#1MS, Q=> TON3_State); //Set2 dir2
TON4(IN:= MW2.9, PT:= T#1MS, Q=> TON4_State); //Set3 dir1
TON5(IN:= NOT(MW2.9), PT:= T#1MS, Q=> TON5_State); //Set3 dir2
IF NOT(MW2.4) THEN MF1_CW:= FALSE; MF1_CCW:= FALSE; ELSE IF MW2.5 THEN MF1_CW:= FALSE; MF1_CCW:= TON0_State; ELSE MF1_CCW:= FALSE; MF1_CW:= TON1_State; END_IF END_IF //WF1
IF NOT(MW2.6) THEN MF2_CW:= FALSE; MF2_CCW:= FALSE; ELSE IF MW2.7 THEN MF2_CW:= FALSE; MF2_CCW:= TON2_State; ELSE MF2_CCW:= FALSE; MF2_CW:= TON3_State; END_IF END_IF //WF2
IF NOT(MW2.8) THEN MF3_CW:= FALSE; MF3_CCW:= FALSE; ELSE IF MW2.9 THEN MF3_CW:= FALSE; MF3_CCW:= TON4_State; ELSE MF3_CCW:= FALSE; MF3_CW:= TON5_State; END_IF END_IF //WF3
 //Wire feeders speed
//Wire feeders//
//PLASMA//
SetCurrent:= SetCurrent_HMI_Man; //Current set
IF NOT(MW0.7) THEN 
	StartParc:= MW2.0; 
	CMT_PS:= MW2.14; //CMT arc
	IF NOT(PilotArc) THEN IF NOT(MW2.1) THEN MW4.4 := TRUE; ELSE MW4.4 := FALSE; END_IF ELSE MW4.4 := FALSE; END_IF
	StartMArc:= MW2.1; //Main arc	
	MW4.2 := FALSE; MW4.6 := FALSE; 
END_IF//Pilot arc 

//PLASMA//
//CMT//
TON_CMT(IN:= CMT_PlusI OR CMT_MinusI, PT:= T#100MS, Q=> TON_CMT_State); //Таймер імпульсу для зміни значення
TON_CMT1(IN:= NOT(CMT_PlusI) AND NOT(CMT_MinusI), PT:= T#100MS, Q=> TON_CMT_State1); //Таймер паузи для зміни значення
IF SetCurrentCMT_HMI <> PrevCurrentCMT_HMI THEN Counter:= WORD_TO_INT(SetCurrentCMT_HMI) -  WORD_TO_INT(PrevCurrentCMT_HMI); //рахуємо кількість імпульсів
	IF Counter > 0 THEN  //Якщо потрібно збільшувати струм
		IF TON_CMT_State1 THEN CMT_PlusI:= TRUE; END_IF //Імпульс
		IF TON_CMT_State THEN CMT_PlusI:= FALSE; PrevCurrentCMT_HMI:= PrevCurrentCMT_HMI +1; Counter:= Counter -1; END_IF //Пауза + інкремент
	ELSIF Counter < 0 THEN  //Якщо потрібно зменшувати струм
		IF TON_CMT_State1 THEN CMT_MinusI:= TRUE; END_IF  //Імпульс
		IF TON_CMT_State THEN CMT_MinusI:= FALSE; PrevCurrentCMT_HMI:= PrevCurrentCMT_HMI -1; Counter:= Counter +1; END_IF //Пауза + декремент
	END_IF
	ELSE CMT_PlusI:= FALSE; CMT_MinusI:= FALSE; //Вимкнення інкрементального та декрементального реле по дефолту
END_IF
//CMT//


IF MW0.8 OR MW0.9 OR MW0.10 OR MW0.11 OR MW0.12 OR MW0.13 OR MW0.14 OR MW0.15 OR MW2.0 OR MW2.1 OR MW2.2 OR MW2.4 OR MW2.6 OR MW2.8 OR MW2.10 OR MW2.11 OR MW2.12 OR MW2.13 OR MW2.14 THEN
	MW6.14 := TRUE;
ELSE
	MW6.14 := FALSE;
END_IF

ProcON:= MW6.15; //Видача ProcON на робот

END_PROGRAM

// Controller_2A1/Application/Alarms_auto
PROGRAM Alarms_auto
VAR
	TON0: TON;
	TON1: TON;
	TON_Analysys_Pilot: TON;
	TON_Analysys_Main: TON;
	TON_Delay_Stop_PF: TON;
	TON_Delay_Stop_WF: TON;
	TON_Delay_Stop_Emagnet: TON;
	TON_Finish_blow: TON;
	Allow_finish_blow: BOOL;
	Prev_Process: WORD;
	T: BOOL;
	TRIG_MW6_9: BOOL;
END_VAR

TON0(IN:= (Process_Auto = 3 AND Alarms = 0), PT:= WORD_TO_TIME(Check_Voltage_Current_Delay)); //Затримка аналізу Voltage та Current
TON_Analysys_Pilot(IN:= StartParc, PT:= WORD_TO_TIME(Delay_Analysys_Pilot*10));//Затримка аналізу чергової дуги
TON_Analysys_Main(IN:= StartMArc, PT:= WORD_TO_TIME(Delay_Analysys_Main*10));//Затримка аналізу основної дуги

//Аналіз чергової та основної дуги
IF TON_Analysys_Pilot.Q AND NOT(PilotArc) AND Auto_Button_State = 1 THEN MW6.10 := TRUE; IF Alarms = 0 THEN Alarms := 4; END_IF END_IF
IF TON_Analysys_Main.Q AND NOT(MainArc) AND Auto_Button_State = 1 THEN MW6.10 := TRUE; IF Alarms = 0 THEN Alarms := 5; END_IF END_IF

//Check Voltage and Current
IF TON0.Q THEN
	IF Set_Emergency_Voltage > MeasureU AND MW4.0 AND MW4.15 THEN MW6.10 := TRUE; IF Alarms = 0 THEN Alarms := 1; END_IF END_IF
	IF Set_Emergency_Current > MeasureI AND MW4.1 AND MW4.15 THEN MW6.10 := TRUE; IF Alarms = 0 THEN Alarms := 2; END_IF END_IF
END_IF

// Ввікнення аварії при нажатій кнопці Emergency stop
IF NOT(EmergencyExt) AND Process_Auto <> 0 AND Auto_Button_State <> 0 THEN IF Alarms = 0 THEN Alarms := 3;  END_IF  END_IF

//Ready total
IF MW6.0 OR MW4.15 THEN
	IF ((((Auto_Button_State = 1 OR Auto_Button_State = 2) AND (Y1 OR Y2 OR Y3 OR Y4)) OR (Auto_Button_State = 0 AND (MW6.1 OR MW6.2 OR MW6.3 OR MW6.4))) AND 
	EmergencyExt AND NOT(MW6.10) AND Alarms = 0) THEN 
		IF NOT(MW4.3) THEN
			MW6.11 := TRUE;
			//MW0.2
		ELSIF MW4.3 AND MW0.2 THEN
			MW6.11 := TRUE;
		ELSE 
			MW6.11 := FALSE; 
		END_IF
	ELSE 
		MW6.11 := FALSE; 
	END_IF
ELSE
	MW6.11 := FALSE;
END_IF

//Robot not ready
IF MW4.3 AND Auto_Button_State = 1 AND NOT(MW0.2) THEN MW6.10 := TRUE; IF Alarms = 0 THEN Alarms := 6; END_IF END_IF

TON1(IN:= MW6.10, PT:= WORD_TO_TIME(Emergency_Delay)); //Затримка аварійного вимкнення

//Аварійна зупинка
IF (TON1.Q OR Auto_Button_State = 2) AND EmergencyExt THEN
	//YES
	MW6.12 := FALSE;
	
	//Block start
	MW6.6 := TRUE;
	
	//Set stop to button
	IF Auto_Button_State <> 0 THEN Auto_Button_State := 2; END_IF
	
	//Save stop process
	IF Process_Auto <> 6 AND Process_Auto <> 4 THEN Prev_Process := Process_Auto; END_IF
	
	//Pre-blowing
	IF Prev_Process = 1 THEN
		Allow_finish_blow := TRUE;
		
	//Waiting Pilot Arc
	ELSIF Prev_Process = 2 THEN
		//Turn off Pilot Arc
		StartParc:= FALSE;
		Allow_finish_blow := TRUE;
		
	//Working Process and CMT Start
	ELSIF Prev_Process = 3 THEN
		// CMT OFF
		CMT_PS := FALSE;
		CMT_PlusI:= FALSE; CMT_MinusI:= FALSE;
		//Turn off Main Arc
		StartMArc:= FALSE;	
		//Turn off Pilot Arc
		StartParc:= FALSE;
		TON_Delay_Stop_PF(IN:=TON_Delay_Start_PF.Q, PT:=WORD_TO_TIME(Delay_Stop_PF));
		TON_Delay_Stop_WF(IN:=TON_Delay_Start_WF.Q, PT:=WORD_TO_TIME(Delay_Stop_WF));
		TON_Delay_Stop_Emagnet(IN:=TON_Delay_Start_Emagnet.Q, PT:=WORD_TO_TIME(Delay_Stop_Emagnet));
		IF (
			(NOT(MW4.7 OR MW4.8 OR MW4.9 OR MW4.10) OR (((MW4.7 OR MW4.8 OR MW4.9 OR MW4.10) AND NOT(TON_Delay_Start_PF.Q)) OR TON_Delay_Stop_PF.Q)) AND
			(NOT(MW4.12 OR MW4.13 OR MW4.14) OR (((MW4.12 OR MW4.13 OR MW4.14) AND NOT(TON_Delay_Start_WF.Q)) OR TON_Delay_Stop_WF.Q))AND
			(NOT(MW4.11) OR ((MW4.11 AND NOT(TON_Delay_Start_Emagnet.Q)) OR TON_Delay_Stop_Emagnet.Q)) 
			) THEN
				Allow_finish_blow := TRUE;
		ELSE
			Process_Auto := 6;
		END_IF
		
	//Waiting Main Arc
	ELSIF Prev_Process = 8 THEN
		//Turn off Main Arc
		StartMArc:= FALSE;
		//Turn off Pilot Arc
		StartParc:= FALSE;
		Allow_finish_blow := TRUE;
		
	//Waiting Additional equipment
	ELSIF Prev_Process = 9 THEN
		// CMT OFF
		CMT_PS := FALSE;
		CMT_PlusI:= FALSE; CMT_MinusI:= FALSE;
		//Turn off Main Arc
		StartMArc:= FALSE;	
		//Turn off Pilot Arc
		StartParc:= FALSE;
		TON_Delay_Stop_PF(IN:=TON_Delay_Start_PF.Q, PT:=WORD_TO_TIME(Delay_Stop_PF));
		TON_Delay_Stop_WF(IN:=TON_Delay_Start_WF.Q, PT:=WORD_TO_TIME(Delay_Stop_WF));
		TON_Delay_Stop_Emagnet(IN:=TON_Delay_Start_Emagnet.Q, PT:=WORD_TO_TIME(Delay_Stop_Emagnet));
		IF (
			(NOT(MW4.7 OR MW4.8 OR MW4.9 OR MW4.10) OR (((MW4.7 OR MW4.8 OR MW4.9 OR MW4.10) AND NOT(TON_Delay_Start_PF.Q)) OR TON_Delay_Stop_PF.Q)) AND
			(NOT(MW4.12 OR MW4.13 OR MW4.14) OR (((MW4.12 OR MW4.13 OR MW4.14) AND NOT(TON_Delay_Start_WF.Q)) OR TON_Delay_Stop_WF.Q)) AND
			(NOT(MW4.11) OR ((MW4.11 AND NOT(TON_Delay_Start_Emagnet.Q)) OR TON_Delay_Stop_Emagnet.Q))
			) THEN
				Allow_finish_blow := TRUE;
		ELSE
			Process_Auto := 6;
		END_IF
	END_IF
	IF TON_Delay_Stop_PF.Q THEN PF1 := FALSE; PF2 := FALSE; PF3 := FALSE; PF4 := FALSE; Y5 := FALSE; Y6 := FALSE; Y7 := FALSE; Y8 := FALSE; END_IF
	IF TON_Delay_Stop_WF.Q THEN MF1_CW:= FALSE; MF1_CCW := FALSE; MF2_CW:= FALSE; MF2_CCW := FALSE; MF3_CW:= FALSE; MF3_CCW := FALSE; END_IF
	IF (MW4.11 AND NOT(TON_Delay_Start_Emagnet.Q)) OR TON_Delay_Stop_Emagnet.Q OR Allow_finish_blow THEN 
		//Вимикаємо магніт
		EM_R_EN := FALSE;
		EM_L_EN := FALSE;
		EM_R_PWM := FALSE;
		EM_L_PWM := FALSE;
		ToggleState := FALSE;
		LastToggleTime := 0;
	ELSIF Prev_Process <> 1 AND Prev_Process <> 2 AND Prev_Process <> 8 AND Auto_Button_State <> 0 AND Prev_Process <> 0 THEN
		IF MW4.11 THEN
				EM_R_EN := TRUE;
				EM_L_EN := TRUE;
				HalfPeriod_us := REAL_TO_ULINT(1000000.0 / EmagFreqCalc_Auto / 2.0); //Період в мікросекундах
				SysTimeGetUs(CurrentTime); // CurrentTime ULINT
				IF (CurrentTime - LastToggleTime) >= HalfPeriod_us THEN //Перевірка пройденого часу
					ToggleState := NOT(ToggleState); //Інверсія
					LastToggleTime := CurrentTime; //Обнулення таймеру
				END_IF	
				EM_R_PWM := ToggleState;
				EM_L_PWM := NOT(ToggleState);
		END_IF
	END_IF
	//Finish blowing
	IF Allow_finish_blow THEN
				TON_Finish_blow(IN:=Enable_Start, PT:=WORD_TO_TIME(Delay_Gas_Finishblow * 10));
				//Finish blow
				IF TON_Finish_blow.Q THEN Allow_finish_blow := FALSE; Y1 := FALSE; Y2 := FALSE; Y3 := FALSE; Y4 := FALSE; Enable_Start := FALSE; Process_Auto := 0; 
				TON_Delay_Stop_PF(IN:=FALSE); TON_Delay_Stop_Emagnet(IN:=FALSE); TON_Delay_Stop_WF(IN:=FALSE); TON_Finish_blow(IN:=FALSE);
				TON_Delay_Start_PF(IN:=FALSE); TON_Delay_Start_Emagnet(IN:=FALSE); TON_Delay_Start_WF(IN:=FALSE);TON_preblow(IN:=FALSE);
				MW6.13 := FALSE;
				Auto_Button_State := 0;
				Prev_Process := 0;
				ELSE Process_Auto := 4; END_IF
				
	END_IF
ELSIF NOT(TON1.Q) AND MW6.10 THEN
	IF MW4.11 THEN
				EM_R_EN := TRUE;
				EM_L_EN := TRUE;
				HalfPeriod_us := REAL_TO_ULINT(1000000.0 / EmagFreqCalc_Auto / 2.0); //Період в мікросекундах
				SysTimeGetUs(CurrentTime); // CurrentTime ULINT
				IF (CurrentTime - LastToggleTime) >= HalfPeriod_us THEN //Перевірка пройденого часу
					ToggleState := NOT(ToggleState); //Інверсія
					LastToggleTime := CurrentTime; //Обнулення таймеру
				END_IF	
				EM_R_PWM := ToggleState;
				EM_L_PWM := NOT(ToggleState);
	END_IF
END_IF

//Emergency Stop
IF (NOT(EmergencyExt) OR (Process_Auto = 4 OR Process_Auto = 6)) AND Auto_Button_State <> 0 AND NOT(MW6.11) AND Alarms = 3 THEN
	//YES
	MW6.12 := FALSE;
	
	//Block start
	MW6.6 := TRUE;
	
	//Set stop to button
	IF Auto_Button_State <> 0 THEN Auto_Button_State := 2; END_IF
	
	// CMT OFF
	CMT_PS := FALSE;
	CMT_PlusI:= FALSE; CMT_MinusI:= FALSE;
	
	//Turn off Main Arc
	StartMArc:= FALSE;	
	
	//Turn off Pilot Arc
	StartParc:= FALSE;
	
	//Вимикаємо магніт
	EM_R_EN := FALSE;
	EM_L_EN := FALSE;
	EM_R_PWM := FALSE;
	EM_L_PWM := FALSE;
	ToggleState := FALSE;
	LastToggleTime := 0;
	PF1 := FALSE; PF2 := FALSE; PF3 := FALSE; PF4 := FALSE; Y5 := FALSE; Y6 := FALSE; Y7 := FALSE; Y8 := FALSE;
	MF1_CW:= FALSE; MF1_CCW := FALSE; MF2_CW:= FALSE; MF2_CCW := FALSE; MF3_CW:= FALSE; MF3_CCW := FALSE;
	
	//Finish blow
	TON_Finish_blow(IN:=Enable_Start, PT:=WORD_TO_TIME(Delay_Gas_Finishblow * 10));
	IF TON_Finish_blow.Q THEN Allow_finish_blow := FALSE; Y1 := FALSE; Y2 := FALSE; Y3 := FALSE; Y4 := FALSE; Enable_Start := FALSE; Process_Auto := 0; 
		TON_Delay_Stop_PF(IN:=FALSE); TON_Delay_Stop_Emagnet(IN:=FALSE); TON_Delay_Stop_WF(IN:=FALSE); TON_Finish_blow(IN:=FALSE);
		TON_Delay_Start_PF(IN:=FALSE); TON_Delay_Start_Emagnet(IN:=FALSE); TON_Delay_Start_WF(IN:=FALSE);TON_preblow(IN:=FALSE);
		MW6.13 := FALSE;
		Auto_Button_State := 0;
		Prev_Process := 0;
	ELSE Process_Auto := 4; END_IF
END_IF

//Reset Alarm
IF MW4.5 AND Auto_Button_State <> 2 THEN Alarms := 0; MW6.10 := FALSE; MW6.13 := FALSE; MW6.9 := FALSE; MW6.5:= FALSE;  TON_Finish_blow(IN:=FALSE); END_IF //Скидання аларму

END_PROGRAM

// Controller_2A1/Application/Alarms_manual
PROGRAM Alarms_manual
VAR
	TON0: TON;
	TON0_State: BOOL;
	TON2: TON;
	TON1: TON;
	TON_Emergency_Man: BOOL;
	TON3: TON;
END_VAR

TON0(IN:= MW2.0, PT:= WORD_TO_TIME(Check_Voltage_Current_Delay), Q=> TON0_State); //Затримка аналізу аварій

TON2(IN:=  ErrorInManual = 11, PT:= T#1000MS); //Таймер блимання помилки
TON3(IN:=  ErrorInManual = 10, PT:= T#1000MS); //Таймер блимання помилки
IF NOT(MW0.7) THEN ErrorInManual:= 11;
	ELSIF ErrorInManual = 11 AND TON2.Q THEN ErrorInManual:= 10; //Перемикання блималки
	ELSIF ErrorInManual = 10 AND TON3.Q THEN ErrorInManual:= 11; //Перемикання блималки
END_IF

IF TON0_State THEN
	IF Set_Emergency_Voltage > MeasureU AND MW4.0 THEN MW0.7 := TRUE; Alarms := 1; END_IF
	IF Set_Emergency_Current > MeasureI AND MW4.1 THEN MW0.7 := TRUE; Alarms := 2; END_IF
END_IF

IF NOT(MW0.7) AND EmergencyExt AND Alarms = 0 THEN MW0.6 := TRUE; ELSE MW0.6 := FALSE; END_IF//Готовність

IF MW0.7 OR NOT(EmergencyExt) THEN MW0.6 := FALSE; END_IF // Скидання готовності

IF MW0.7 AND Alarms = 0 AND EmergencyExt THEN MW0.7 := FALSE; END_IF
IF NOT(EmergencyExt) THEN Alarms := 3; MW0.7 := TRUE; END_IF // Ввікнення аварії при нажатій кнопці Emergency stop

TON1(IN:= MW0.7 OR NOT(EmergencyExt), PT:= WORD_TO_TIME(Emergency_Delay), Q=> TON_Emergency_Man); //Затримка аварійного вимкнення

//Аварійна зупинка
IF TON_Emergency_Man THEN MW4.2 := TRUE; MW4.4 := TRUE; MW4.6 := TRUE; MW2.0 := FALSE; MW2.1 := FALSE; MW2.10 := FALSE; MW2.11 := FALSE; MW2.12 := FALSE; MW2.13 := FALSE; MW2.4 := FALSE; MW2.6 := FALSE; MW2.8 := FALSE; MW2.2 := FALSE; MW2.14 := FALSE; END_IF

IF MW4.5 THEN Alarms := 0; MW0.7 := FALSE; END_IF //Скидання аларму

END_PROGRAM
